Fanuc KAREL source: KA00155.KL

PROGRAM KA00155
%NOLOCKGROUP
VAR
  SRC: ARRAY[4] OF REAL
  DST: ARRAY[4] OF REAL
BEGIN
  DST = SRC
END KA00155
